Fanuc KAREL source: KA00130.KL

PROGRAM KA00130
%NOLOCKGROUP
VAR
  SRC: ARRAY[2] OF BYTE
  DST: CONFIG
BEGIN
  SRC[1] = 2
  DST = SRC[1]
END KA00130
